(* PLC project zarechnaya.project, CODESYS CODESYS V3.5 SP17 Patch 3 *)
(* stored: creationDateTime 2026-10-20T05:42:22.1876153, modificationDateTime 1601-01-01T03:00:00 *)

(* FB_TimeIdioms — таймеры промывочного насоса (ST, FUNCTION_BLOCK). Поведение (модель scenarios/reference/model_FB_TimeIdioms.py): - fbPulse(IN := NOT fbPulse.Q, PT := T#500MS) — самосбрасывающийся таймер: Q = TRUE ровно на один вызов, когда ET ≥ 500 мс, следующий вызов сбрасывает таймер (IN = FALSE), ещё следующий — запускает снова; xPulse := fbPulse.Q (C2S7-SEM-TIMER-Q: S7-1200 обновляет Q и при чтении члена); - xEarly := fbDelay.Q до вызова fbDelay — значение прошлого вызова; xLate := fbDelay.Q после вызова fbDelay(IN := xIn, PT := T#1S) — TON: Q, когда xIn держится ≥ 1 с; - xLong := tIn > T#30D — литерал больше диапазона Time S7 (±24d20h): на S7-1500 → LTime, на S7-1200 — impossible (C2S7-TYPE-TIME). TIME CODESYS — 32 бита без знака. *)
FUNCTION_BLOCK FB_TimeIdioms
  VAR_INPUT
    xIn : BOOL;
    tIn : TIME;
  END_VAR
  VAR_OUTPUT
    xPulse : BOOL;
    xEarly : BOOL;
    xLate : BOOL;
    xLong : BOOL;
  END_VAR
  VAR
    fbPulse : TON;
    fbDelay : TON;
  END_VAR

            fbPulse(IN := NOT fbPulse.Q, PT := T#500MS);
xPulse := fbPulse.Q;
xEarly := fbDelay.Q;
fbDelay(IN := xIn, PT := T#1S);
xLate := fbDelay.Q;
xLong := tIn > T#30D;

          
END_FUNCTION_BLOCK
